Fanuc KAREL source: kb00112.KL

PROGRAM KB00112
%STACKSIZE=65535
%PRIORITY=65535
%NOLOCKGROUP
VAR
P1 : JOINTPOS9
RESULT : BOOLEAN
BEGIN
-- UNRESOLVED_PC line 7 opcodes [27 22 1C 27 9D 76 23] marker_code=0
END KB00112
